Fanuc KAREL source: KB00045.KL

PROGRAM KB00045
%NOLOCKGROUP
%ENVIRONMENT MULTI
VAR
  P1: STRING[80]
  P2: INTEGER
BEGIN
  P1 = 'A'
  P2 = 1
  CONT_TASK(P1, P2)
END KB00045
